{region 'Documentation'}
(*!
<summary>Returns whole calendar days since 1970-01-01; ignores any time-of-day remainder.</summary>
*)
{endregion}
FUNCTION INTERNAL DateToDayNumber : UDINT //! Whole days since 1970-01-01.
VAR_INPUT
    Value : DATE; //! Calendar date; any stored time-of-day remainder is ignored.
END_VAR
VAR CONSTANT
    SecondsPerDay : UDINT := 86400;
END_VAR

DateToDayNumber := DATE_TO_UDINT(Value) / SecondsPerDay;

END_FUNCTION

(* stored: Version 1.1.0.1
   POU DateToDayNumber: Id {0cd4f77c-e986-444a-8053-ecade3357c1d}, SpecialFunc None *)
